// Réception des alarmes (docs/04 § 4, docs/14)
INTERFACE I_AlarmSink

METHOD Raise
VAR_INPUT
    nGlobalId : UDINT;
    nCode : UINT;
    nSubCode : UDINT;
    eSeverity : E_Severity;
END_VAR
END_METHOD

METHOD Clear
VAR_INPUT
    nGlobalId : UDINT;
    nCode : UINT;
END_VAR
END_METHOD

END_INTERFACE

(* stored: Version 1.1.0.1, ProductVersion 3.1.4024.12
   Itf I_AlarmSink: Id {f97f1660-5141-5b18-bf2e-5411ee34d188}
   Method Raise: Id {7acab48b-09b7-5727-88b6-c5c775cd2aa4}
   Method Clear: Id {9d337b43-f468-5a49-9c75-738e489f980f} *)
